// TIA Portal V21 export
// export: Created 2026-10-23T20:44:46.9310721Z, ExportSetting WithDefaults, DisplayName Totally Integrated Automation Portal, DisplayVersion V21 Update 1, DisplayName SINAMICS Startdrive Advanced, DisplayVersion V21 HF2, DisplayName SINAMICS Startdrive G110M, G120, G120C, G120D, G120P, G115D, DisplayVersion V21 HF2, DisplayName SINAMICS Startdrive G130, G150, S120, S150, G200, G220, S200, S210, S220, Innomotics MVD, DisplayVersion V21 HF2, DisplayName STEP 7 Professional, DisplayVersion V21 Update 1, DisplayName STEP 7 Safety, DisplayVersion V21, DisplayName Tech WebApplication, DisplayVersion V21, DisplayName WinCC Basic/Comfort/Advanced, DisplayVersion V21 Update 1, DisplayName WinCC Unified, DisplayVersion V21 Update 1
ORGANIZATION_BLOCK "OB_Main"   // OB1, SCL, ProgramCycle
TITLE = "Main Program Sweep (Cycle)" / Main program of PLC_1200
{ S7_Optimized_Access := 'TRUE' }
VERSION : 0.1
// Calls the conveyor with the onboard inputs and output of the CPU 1214C
// stored: AutoNumber true, IsIECCheckEnabled false, SetENOAutomatically false
   VAR_INPUT
      Initial_Call : Bool;   // Initial call of this OB
      Remanence : Bool;   // =True, if remanent data are available
   END_VAR
BEGIN

       REGION Conveyor
           "IDB_Conveyor1200"(Start := "BeltStart",
                              Stop := "BeltStop",
                              SpeedRaw := "BeltSpeedRaw",
                              Motor => "BeltMotor");
       END_REGION
END_ORGANIZATION_BLOCK
